// SIMATIC S7-200 project (STEP 7-Micro/WIN), CPU 224 CN REL 02.01

SYMBOL_TABLE Usuario 1
Run              M10.0
Sensor_base      I0.0
X_limite_adelante I0.1
X_limite_atras   I0.2
Y_limite_adelante I0.3
Y_limite_atras   I0.4
Switch           I0.5
Reset            I0.6
Start_y_s1       I0.7
Boton_stop_y_s2  I1.0
Boton_s3_derecha I1.1
Boton_s4_adelante I1.2
Boton_s5_atras   I1.3
Boton_s6_arriba  I1.4
Boton_s7_abajo   I1.5
Pulso_en_Z       Q0.0
Pulso_en_XY      Q0.1
Dir_Eje_Z        Q0.2
Dir_eje_X        Q0.3
Dir_Eje_Y        Q0.4
Pulso_en_X       Q0.5
Pulso_en_Y       Q0.6
Pinza            Q0.7
Posicion_de_Z    VD210
Posicion_de_XY   VD220
Posicion_de_X    VD230
Posicion_de_Y    VD240
Velocidad_de_Z   VD250
Velocidad_de_XY  VD260
END_SYMBOL_TABLE

ORGANIZATION_BLOCK Principal:OB1
TITLE=Notas del programa
BEGIN
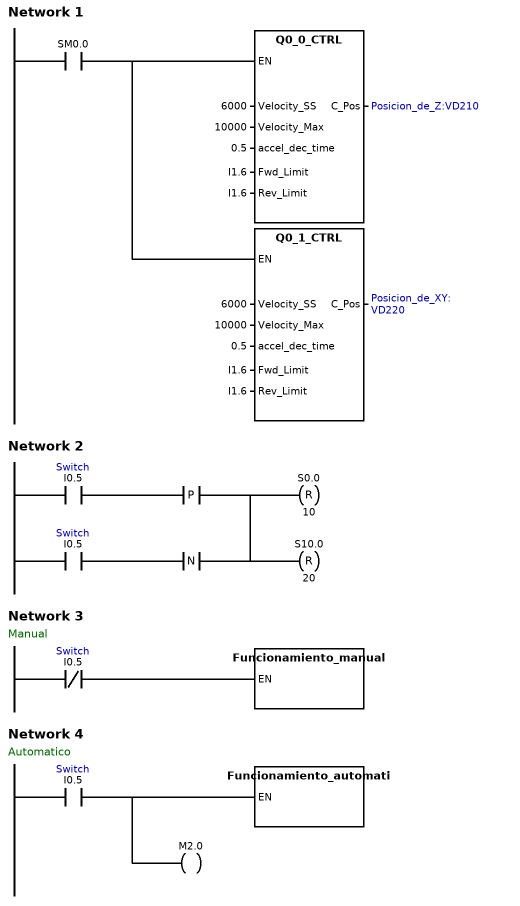
Network 1
// (network saved uncompiled; LAD cells follow)
// row 0: c0 -| |- SM0.0 v  c1 --  c2 [Q0_0_CTRL EN:=power@row0, Velocity_SS:=6000, Velocity_Max:=10000, accel_dec_time:=0.5, Fwd_Limit:=I1.6, Rev_Limit:=I1.6, C_Pos=>Posicion_de_Z:VD210]
// row 1: c0 ^v  c2 [box]
// row 2: c0 ^v  c2 [box]
// row 3: c0 ^  c1 --  c2 [Q0_1_CTRL EN:=power@row3, Velocity_SS:=6000, Velocity_Max:=10000, accel_dec_time:=0.5, Fwd_Limit:=I1.6, Rev_Limit:=I1.6, C_Pos=>Posicion_de_XY:VD220]
// row 4: c2 [box]
// row 5: c2 [box]
Network 2
// (network saved uncompiled; LAD cells follow)
// row 0: c0 -| |- Switch:I0.5  c1 -|P|-  v  c2 -(R) S0.0, 10
// row 1: c0 -| |- Switch:I0.5  c1 -|N|-  ^  c2 -(R) S10.0, 20
Network 3
// Manual
// (network saved uncompiled; LAD cells follow)
// row 0: c0 -|/|- Switch:I0.5  c1 --  c2 [Funcionamiento_manual EN:=power@row0]
Network 4
// Automatico
// (network saved uncompiled; LAD cells follow)
// row 0: c0 -| |- Switch:I0.5 v  c1 --  c2 [Funcionamiento_automati EN:=power@row0]
// row 1: c0 ^  c1 -( ) M2.0
END_ORGANIZATION_BLOCK

SUBROUTINE_BLOCK Funcionamiento_manual:SBR0
TITLE=
BEGIN
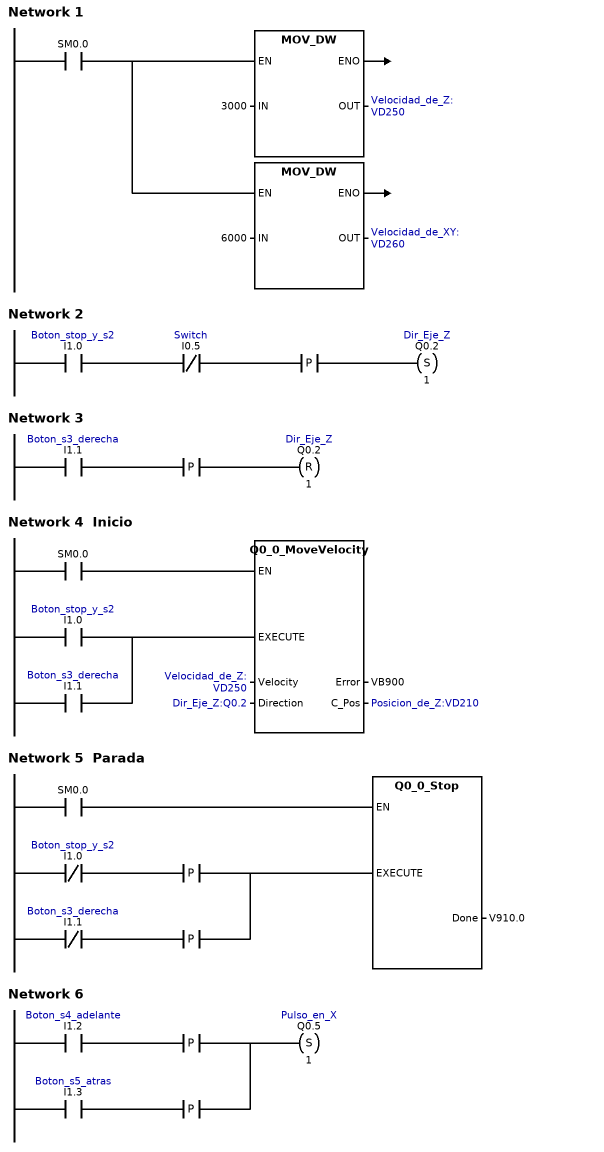
Network 1
// (network saved uncompiled; LAD cells follow)
// row 0: c0 -| |- SM0.0 v  c1 --  c2 [MOV_DW EN:=power@row0, IN:=3000, ENO=>power, OUT=>Velocidad_de_Z:VD250]  c3 ->
// row 1: c0 ^v  c2 [box]
// row 2: c0 ^  c1 --  c2 [MOV_DW EN:=power@row2, IN:=6000, ENO=>power, OUT=>Velocidad_de_XY:VD260]  c3 ->
// row 3: c2 [box]
Network 2
// (network saved uncompiled; LAD cells follow)
// row 0: c0 -| |- Boton_stop_y_s2:I1.0  c1 -|/|- Switch:I0.5  c2 -|P|-  c3 -(S) Dir_Eje_Z:Q0.2, 1
Network 3
// (network saved uncompiled; LAD cells follow)
// row 0: c0 -| |- Boton_s3_derecha:I1.1  c1 -|P|-  c2 -(R) Dir_Eje_Z:Q0.2, 1
Network 4 // Inicio
// (network saved uncompiled; LAD cells follow)
// row 0: c0 -| |- SM0.0  c1 --  c2 [Q0_0_MoveVelocity EN:=power@row0, EXECUTE:=power@row1, Velocity:=Velocidad_de_Z:VD250, Direction:=Dir_Eje_Z:Q0.2, Error=>VB900, C_Pos=>Posicion_de_Z:VD210]
// row 1: c0 -| |- Boton_stop_y_s2:I1.0 v  c1 --  c2 [box]
// row 2: c0 -| |- Boton_s3_derecha:I1.1 ^  c2 [box]
Network 5 // Parada
// (network saved uncompiled; LAD cells follow)
// row 0: c0 -| |- SM0.0  c1 --  c2 --  c3 [Q0_0_Stop EN:=power@row0, EXECUTE:=power@row1, Done=>V910.0]
// row 1: c0 -|/|- Boton_stop_y_s2:I1.0  c1 -|P|-  v  c2 --  c3 [box]
// row 2: c0 -|/|- Boton_s3_derecha:I1.1  c1 -|P|-  ^  c3 [box]
Network 6
// (network saved uncompiled; LAD cells follow)
// row 0: c0 -| |- Boton_s4_adelante:I1.2  c1 -|P|-  v  c2 -(S) Pulso_en_X:Q0.5, 1
// row 1: c0 -| |- Boton_s5_atras:I1.3  c1 -|P|-  ^
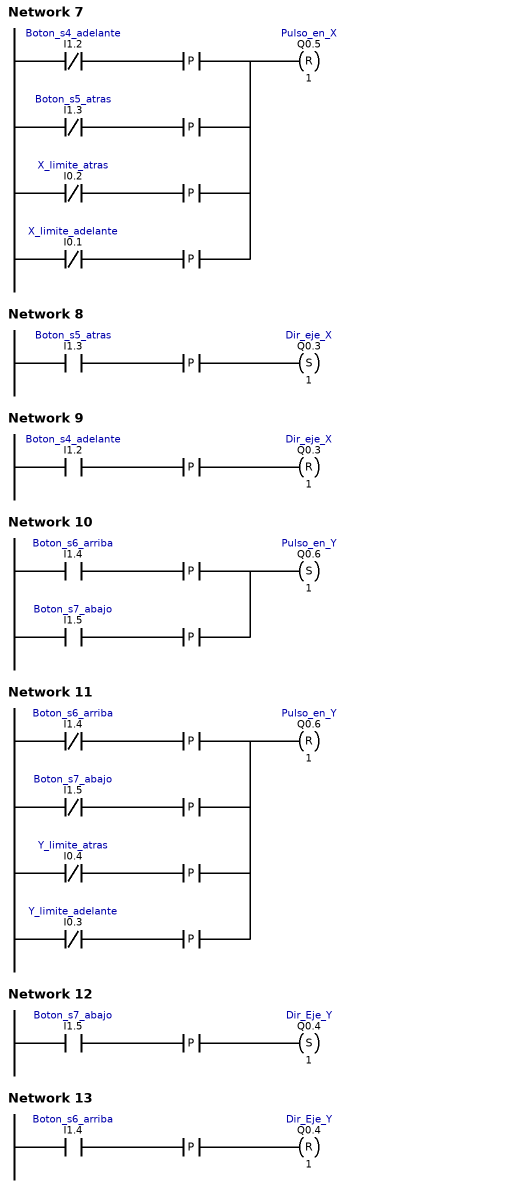
Network 7
// (network saved uncompiled; LAD cells follow)
// row 0: c0 -|/|- Boton_s4_adelante:I1.2  c1 -|P|-  v  c2 -(R) Pulso_en_X:Q0.5, 1
// row 1: c0 -|/|- Boton_s5_atras:I1.3  c1 -|P|-  ^v
// row 2: c0 -|/|- X_limite_atras:I0.2  c1 -|P|-  ^v
// row 3: c0 -|/|- X_limite_adelante:I0.1  c1 -|P|-  ^
Network 8
// (network saved uncompiled; LAD cells follow)
// row 0: c0 -| |- Boton_s5_atras:I1.3  c1 -|P|-  c2 -(S) Dir_eje_X:Q0.3, 1
Network 9
// (network saved uncompiled; LAD cells follow)
// row 0: c0 -| |- Boton_s4_adelante:I1.2  c1 -|P|-  c2 -(R) Dir_eje_X:Q0.3, 1
Network 10
// (network saved uncompiled; LAD cells follow)
// row 0: c0 -| |- Boton_s6_arriba:I1.4  c1 -|P|-  v  c2 -(S) Pulso_en_Y:Q0.6, 1
// row 1: c0 -| |- Boton_s7_abajo:I1.5  c1 -|P|-  ^
Network 11
// (network saved uncompiled; LAD cells follow)
// row 0: c0 -|/|- Boton_s6_arriba:I1.4  c1 -|P|-  v  c2 -(R) Pulso_en_Y:Q0.6, 1
// row 1: c0 -|/|- Boton_s7_abajo:I1.5  c1 -|P|-  ^v
// row 2: c0 -|/|- Y_limite_atras:I0.4  c1 -|P|-  ^v
// row 3: c0 -|/|- Y_limite_adelante:I0.3  c1 -|P|-  ^
Network 12
// (network saved uncompiled; LAD cells follow)
// row 0: c0 -| |- Boton_s7_abajo:I1.5  c1 -|P|-  c2 -(S) Dir_Eje_Y:Q0.4, 1
Network 13
// (network saved uncompiled; LAD cells follow)
// row 0: c0 -| |- Boton_s6_arriba:I1.4  c1 -|P|-  c2 -(R) Dir_Eje_Y:Q0.4, 1
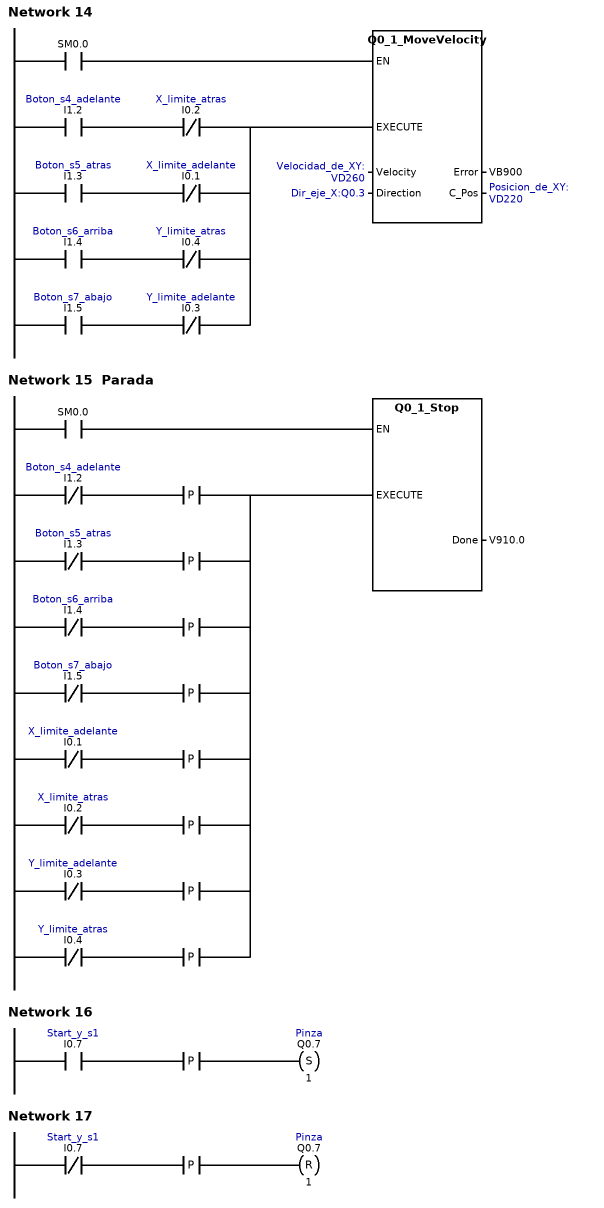
Network 14
// (network saved uncompiled; LAD cells follow)
// row 0: c0 -| |- SM0.0  c1 --  c2 --  c3 [Q0_1_MoveVelocity EN:=power@row0, EXECUTE:=power@row1, Velocity:=Velocidad_de_XY:VD260, Direction:=Dir_eje_X:Q0.3, Error=>VB900, C_Pos=>Posicion_de_XY:VD220]
// row 1: c0 -| |- Boton_s4_adelante:I1.2  c1 -|/|- X_limite_atras:I0.2 v  c2 --  c3 [box]
// row 2: c0 -| |- Boton_s5_atras:I1.3  c1 -|/|- X_limite_adelante:I0.1 ^v  c3 [box]
// row 3: c0 -| |- Boton_s6_arriba:I1.4  c1 -|/|- Y_limite_atras:I0.4 ^v
// row 4: c0 -| |- Boton_s7_abajo:I1.5  c1 -|/|- Y_limite_adelante:I0.3 ^
Network 15 // Parada
// (network saved uncompiled; LAD cells follow)
// row 0: c0 -| |- SM0.0  c1 --  c2 --  c3 [Q0_1_Stop EN:=power@row0, EXECUTE:=power@row1, Done=>V910.0]
// row 1: c0 -|/|- Boton_s4_adelante:I1.2  c1 -|P|-  v  c2 --  c3 [box]
// row 2: c0 -|/|- Boton_s5_atras:I1.3  c1 -|P|-  ^v  c3 [box]
// row 3: c0 -|/|- Boton_s6_arriba:I1.4  c1 -|P|-  ^v
// row 4: c0 -|/|- Boton_s7_abajo:I1.5  c1 -|P|-  ^v
// row 5: c0 -|/|- X_limite_adelante:I0.1  c1 -|P|-  ^v
// row 6: c0 -|/|- X_limite_atras:I0.2  c1 -|P|-  ^v
// row 7: c0 -|/|- Y_limite_adelante:I0.3  c1 -|P|-  ^v
// row 8: c0 -|/|- Y_limite_atras:I0.4  c1 -|P|-  ^
Network 16
// (network saved uncompiled; LAD cells follow)
// row 0: c0 -| |- Start_y_s1:I0.7  c1 -|P|-  c2 -(S) Pinza:Q0.7, 1
Network 17
// (network saved uncompiled; LAD cells follow)
// row 0: c0 -|/|- Start_y_s1:I0.7  c1 -|P|-  c2 -(R) Pinza:Q0.7, 1
Network 22 // 网络标题
// 网络注释
END_SUBROUTINE_BLOCK

// SBR1: protected block, not included

// SBR2: protected block, not included

// SBR3: protected block, not included

// SBR4: protected block, not included

// SBR5: protected block, not included

// SBR6: protected block, not included

SUBROUTINE_BLOCK Origen:SBR7
TITLE=
VAR_INPUT
EXECUTE:BOOL;	// L0.0 
END_VAR
VAR_OUTPUT
Done:BOOL;	// L0.1 
END_VAR
BEGIN
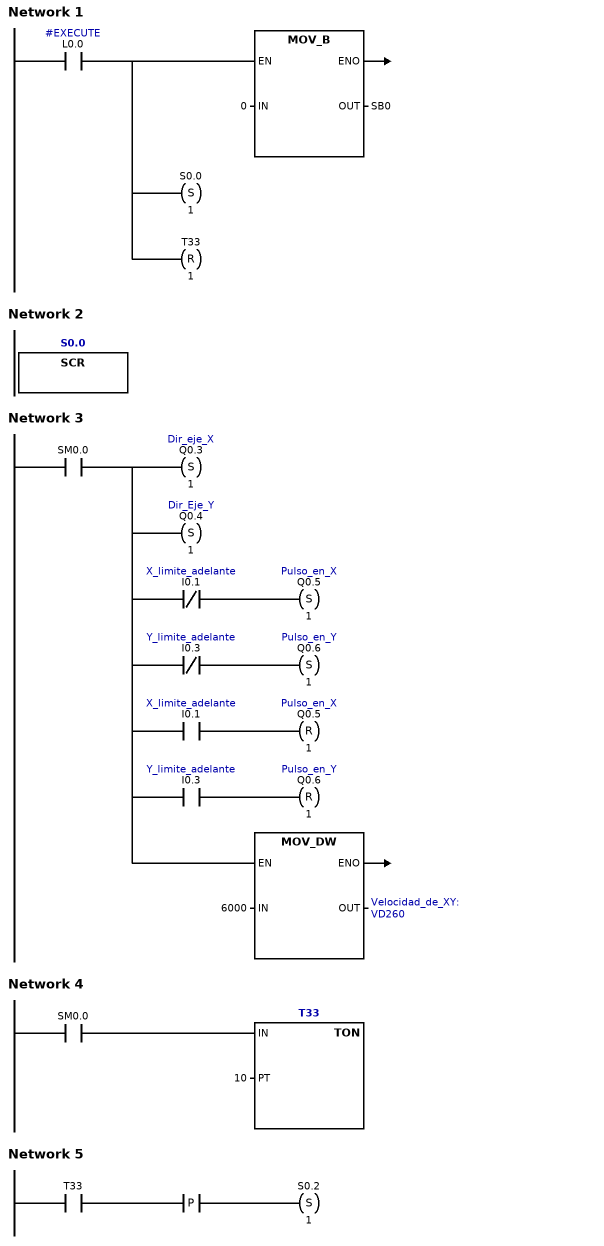
Network 1
LD     #EXECUTE:L0.0
MOVB   0, SB0
S      S0.0, 1
R      T33, 1
Network 2
LSCR   S0.0
Network 3
// (network saved uncompiled; LAD cells follow)
// row 0: c0 -| |- SM0.0 v  c1 -(S) Dir_eje_X:Q0.3, 1
// row 1: c0 ^v  c1 -(S) Dir_Eje_Y:Q0.4, 1
// row 2: c0 ^v  c1 -|/|- X_limite_adelante:I0.1  c2 -(S) Pulso_en_X:Q0.5, 1
// row 3: c0 ^v  c1 -|/|- Y_limite_adelante:I0.3  c2 -(S) Pulso_en_Y:Q0.6, 1
// row 4: c0 ^v  c1 -| |- X_limite_adelante:I0.1  c2 -(R) Pulso_en_X:Q0.5, 1
// row 5: c0 ^v  c1 -| |- Y_limite_adelante:I0.3  c2 -(R) Pulso_en_Y:Q0.6, 1
// row 6: c0 ^  c1 --  c2 [MOV_DW EN:=power@row6, IN:=6000, ENO=>power, OUT=>Velocidad_de_XY:VD260]  c3 ->
// row 7: c2 [box]
Network 4
LD     SM0.0
TON    T33, 10
Network 5
LD     T33
EU
S      S0.2, 1
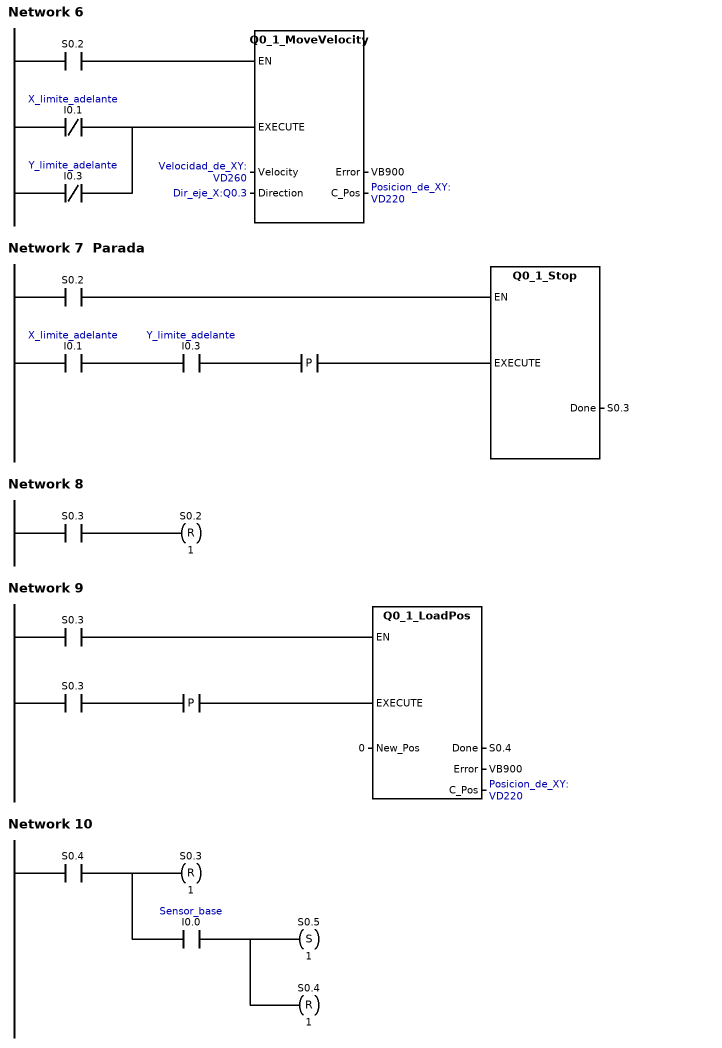
Network 6
// (network saved uncompiled; LAD cells follow)
// row 0: c0 -| |- S0.2  c1 --  c2 [Q0_1_MoveVelocity EN:=power@row0, EXECUTE:=power@row1, Velocity:=Velocidad_de_XY:VD260, Direction:=Dir_eje_X:Q0.3, Error=>VB900, C_Pos=>Posicion_de_XY:VD220]
// row 1: c0 -|/|- X_limite_adelante:I0.1 v  c1 --  c2 [box]
// row 2: c0 -|/|- Y_limite_adelante:I0.3 ^  c2 [box]
Network 7 // Parada
// (network saved uncompiled; LAD cells follow)
// row 0: c0 -| |- S0.2  c1 --  c2 --  c3 --  c4 [Q0_1_Stop EN:=power@row0, EXECUTE:=power@row1, Done=>S0.3]
// row 1: c0 -| |- X_limite_adelante:I0.1  c1 -| |- Y_limite_adelante:I0.3  c2 -|P|-  c3 --  c4 [box]
// row 2: c4 [box]
Network 8
LD     S0.3
R      S0.2, 1
Network 9
// (network saved uncompiled; LAD cells follow)
// row 0: c0 -| |- S0.3  c1 --  c2 --  c3 [Q0_1_LoadPos EN:=power@row0, EXECUTE:=power@row1, New_Pos:=0, Done=>S0.4, Error=>VB900, C_Pos=>Posicion_de_XY:VD220]
// row 1: c0 -| |- S0.3  c1 -|P|-  c2 --  c3 [box]
// row 2: c3 [box]
Network 10
// (network saved uncompiled; LAD cells follow)
// row 0: c0 -| |- S0.4 v  c1 -(R) S0.3, 1
// row 1: c0 ^  c1 -| |- Sensor_base:I0.0 v  c2 -(S) S0.5, 1
// row 2: c1 ^  c2 -(R) S0.4, 1
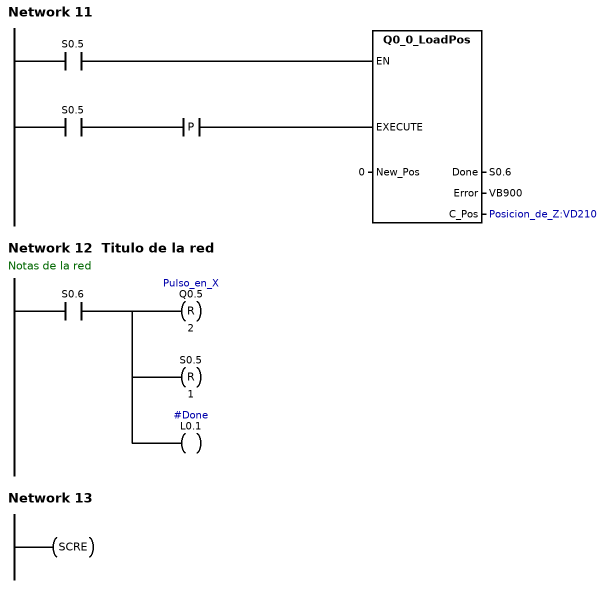
Network 11
// (network saved uncompiled; LAD cells follow)
// row 0: c0 -| |- S0.5  c1 --  c2 --  c3 [Q0_0_LoadPos EN:=power@row0, EXECUTE:=power@row1, New_Pos:=0, Done=>S0.6, Error=>VB900, C_Pos=>Posicion_de_Z:VD210]
// row 1: c0 -| |- S0.5  c1 -|P|-  c2 --  c3 [box]
// row 2: c3 [box]
Network 12 // Titulo de la red
// Notas de la red
// (network saved uncompiled; LAD cells follow)
// row 0: c0 -| |- S0.6 v  c1 -(R) Pulso_en_X:Q0.5, 2
// row 1: c0 ^v  c1 -(R) S0.5, 1
// row 2: c0 ^  c1 -( ) #Done:L0.1
Network 13
SCRE
Network 25 // 网络标题
// 网络注释
END_SUBROUTINE_BLOCK

SUBROUTINE_BLOCK Funcionamiento_automati:SBR8
TITLE=
BEGIN
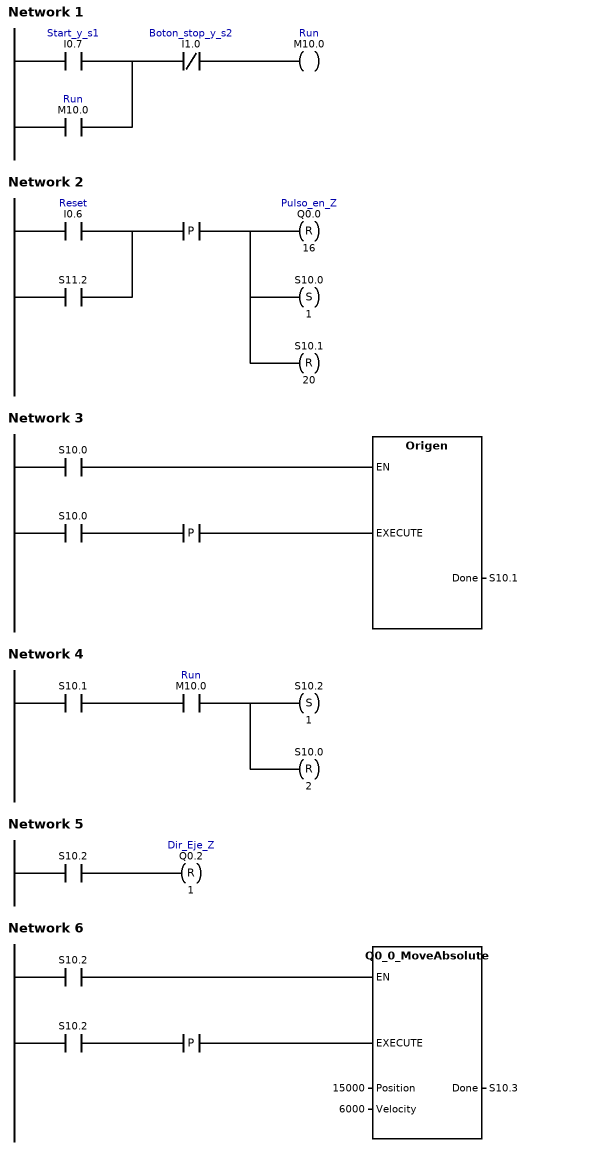
Network 1
// (network saved uncompiled; LAD cells follow)
// row 0: c0 -| |- Start_y_s1:I0.7 v  c1 -|/|- Boton_stop_y_s2:I1.0  c2 -( ) Run:M10.0
// row 1: c0 -| |- Run:M10.0 ^
Network 2
// (network saved uncompiled; LAD cells follow)
// row 0: c0 -| |- Reset:I0.6 v  c1 -|P|-  v  c2 -(R) Pulso_en_Z:Q0.0, 16
// row 1: c0 -| |- S11.2 ^  c1 ^v  c2 -(S) S10.0, 1
// row 2: c1 ^  c2 -(R) S10.1, 20
Network 3
LD     S10.0
=      L60.0
LD     S10.0
EU
=      L63.7
LD     L60.0
CALL   Origen:SBR7, L63.7, S10.1
Network 4
// (network saved uncompiled; LAD cells follow)
// row 0: c0 -| |- S10.1  c1 -| |- Run:M10.0 v  c2 -(S) S10.2, 1
// row 1: c1 ^  c2 -(R) S10.0, 2
Network 5
// (network saved uncompiled; LAD cells follow)
// row 0: c0 -| |- S10.2  c1 -(R) Dir_Eje_Z:Q0.2, 1
Network 6
LD     S10.2
=      L60.0
LD     S10.2
EU
=      L63.7
LD     L60.0
CALL   Q0_0_MoveAbsolute:SBR4, L63.7, 15000, 6000, S10.3
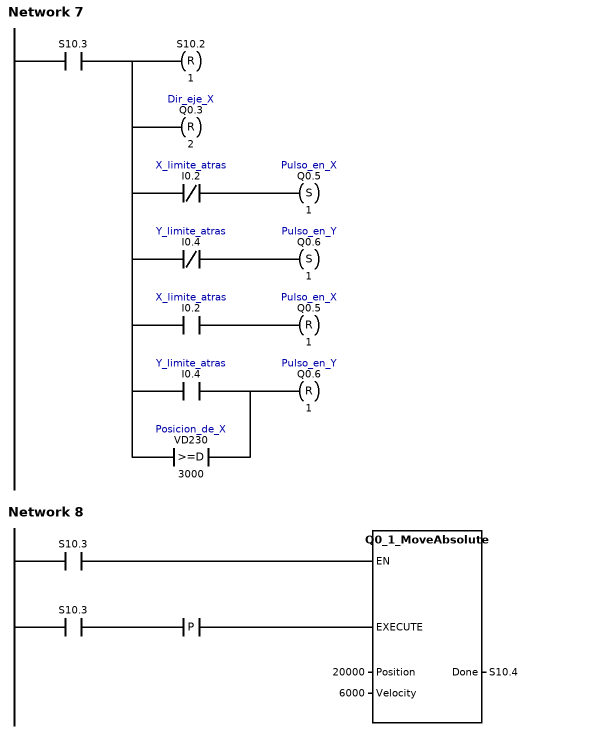
Network 7
// (network saved uncompiled; LAD cells follow)
// row 0: c0 -| |- S10.3 v  c1 -(R) S10.2, 1
// row 1: c0 ^v  c1 -(R) Dir_eje_X:Q0.3, 2
// row 2: c0 ^v  c1 -|/|- X_limite_atras:I0.2  c2 -(S) Pulso_en_X:Q0.5, 1
// row 3: c0 ^v  c1 -|/|- Y_limite_atras:I0.4  c2 -(S) Pulso_en_Y:Q0.6, 1
// row 4: c0 ^v  c1 -| |- X_limite_atras:I0.2  c2 -(R) Pulso_en_X:Q0.5, 1
// row 5: c0 ^v  c1 -| |- Y_limite_atras:I0.4 v  c2 -(R) Pulso_en_Y:Q0.6, 1
// row 6: c0 ^  c1 -|>=D|- Posicion_de_X:VD230, 3000 ^
Network 8
LD     S10.3
=      L60.0
LD     S10.3
EU
=      L63.7
LD     L60.0
CALL   Q0_1_MoveAbsolute:SBR19, L63.7, 20000, 6000, S10.4
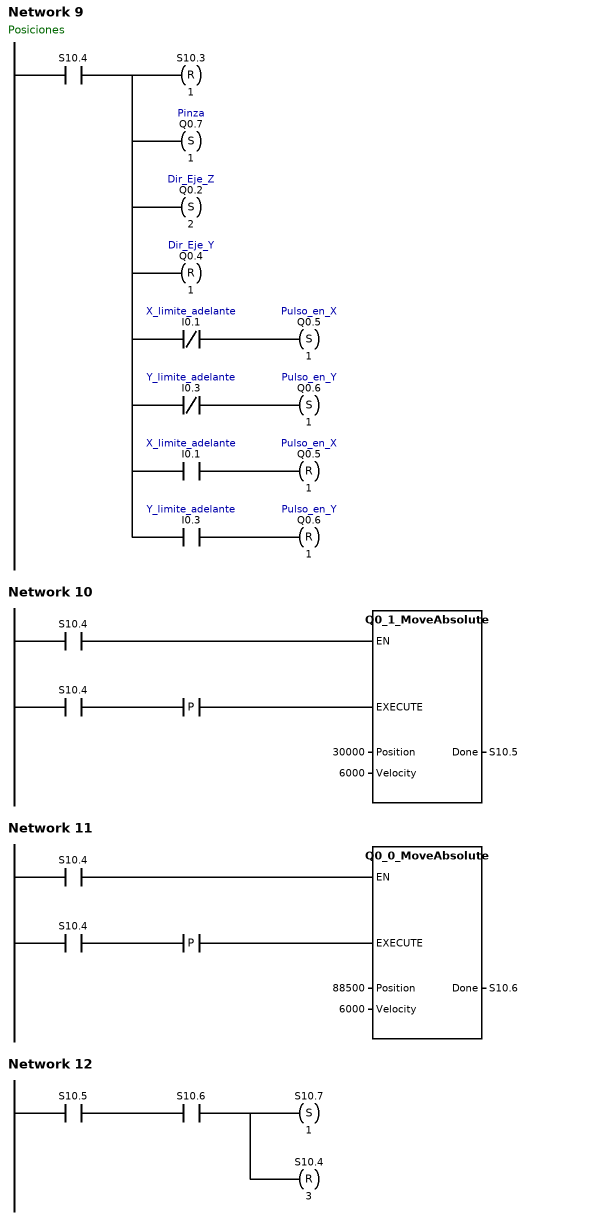
Network 9
// Posiciones
// (network saved uncompiled; LAD cells follow)
// row 0: c0 -| |- S10.4 v  c1 -(R) S10.3, 1
// row 1: c0 ^v  c1 -(S) Pinza:Q0.7, 1
// row 2: c0 ^v  c1 -(S) Dir_Eje_Z:Q0.2, 2
// row 3: c0 ^v  c1 -(R) Dir_Eje_Y:Q0.4, 1
// row 4: c0 ^v  c1 -|/|- X_limite_adelante:I0.1  c2 -(S) Pulso_en_X:Q0.5, 1
// row 5: c0 ^v  c1 -|/|- Y_limite_adelante:I0.3  c2 -(S) Pulso_en_Y:Q0.6, 1
// row 6: c0 ^v  c1 -| |- X_limite_adelante:I0.1  c2 -(R) Pulso_en_X:Q0.5, 1
// row 7: c0 ^  c1 -| |- Y_limite_adelante:I0.3  c2 -(R) Pulso_en_Y:Q0.6, 1
Network 10
LD     S10.4
=      L60.0
LD     S10.4
EU
=      L63.7
LD     L60.0
CALL   Q0_1_MoveAbsolute:SBR19, L63.7, 30000, 6000, S10.5
Network 11
LD     S10.4
=      L60.0
LD     S10.4
EU
=      L63.7
LD     L60.0
CALL   Q0_0_MoveAbsolute:SBR4, L63.7, 88500, 6000, S10.6
Network 12
LD     S10.5
A      S10.6
S      S10.7, 1
R      S10.4, 3
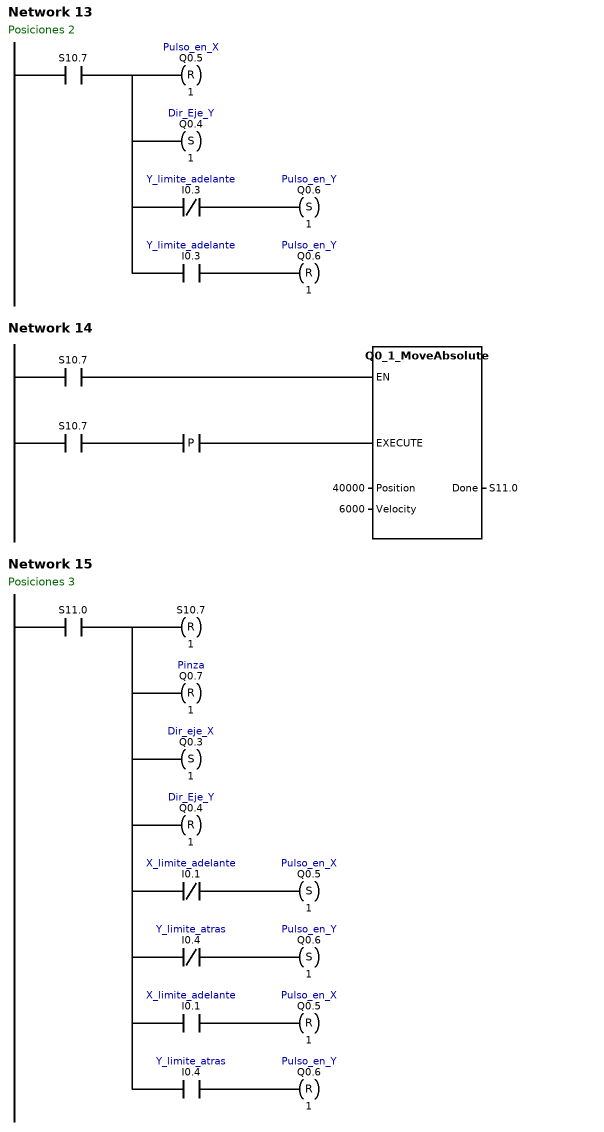
Network 13
// Posiciones 2
// (network saved uncompiled; LAD cells follow)
// row 0: c0 -| |- S10.7 v  c1 -(R) Pulso_en_X:Q0.5, 1
// row 1: c0 ^v  c1 -(S) Dir_Eje_Y:Q0.4, 1
// row 2: c0 ^v  c1 -|/|- Y_limite_adelante:I0.3  c2 -(S) Pulso_en_Y:Q0.6, 1
// row 3: c0 ^  c1 -| |- Y_limite_adelante:I0.3  c2 -(R) Pulso_en_Y:Q0.6, 1
Network 14
LD     S10.7
=      L60.0
LD     S10.7
EU
=      L63.7
LD     L60.0
CALL   Q0_1_MoveAbsolute:SBR19, L63.7, 40000, 6000, S11.0
Network 15
// Posiciones 3
// (network saved uncompiled; LAD cells follow)
// row 0: c0 -| |- S11.0 v  c1 -(R) S10.7, 1
// row 1: c0 ^v  c1 -(R) Pinza:Q0.7, 1
// row 2: c0 ^v  c1 -(S) Dir_eje_X:Q0.3, 1
// row 3: c0 ^v  c1 -(R) Dir_Eje_Y:Q0.4, 1
// row 4: c0 ^v  c1 -|/|- X_limite_adelante:I0.1  c2 -(S) Pulso_en_X:Q0.5, 1
// row 5: c0 ^v  c1 -|/|- Y_limite_atras:I0.4  c2 -(S) Pulso_en_Y:Q0.6, 1
// row 6: c0 ^v  c1 -| |- X_limite_adelante:I0.1  c2 -(R) Pulso_en_X:Q0.5, 1
// row 7: c0 ^  c1 -| |- Y_limite_atras:I0.4  c2 -(R) Pulso_en_Y:Q0.6, 1
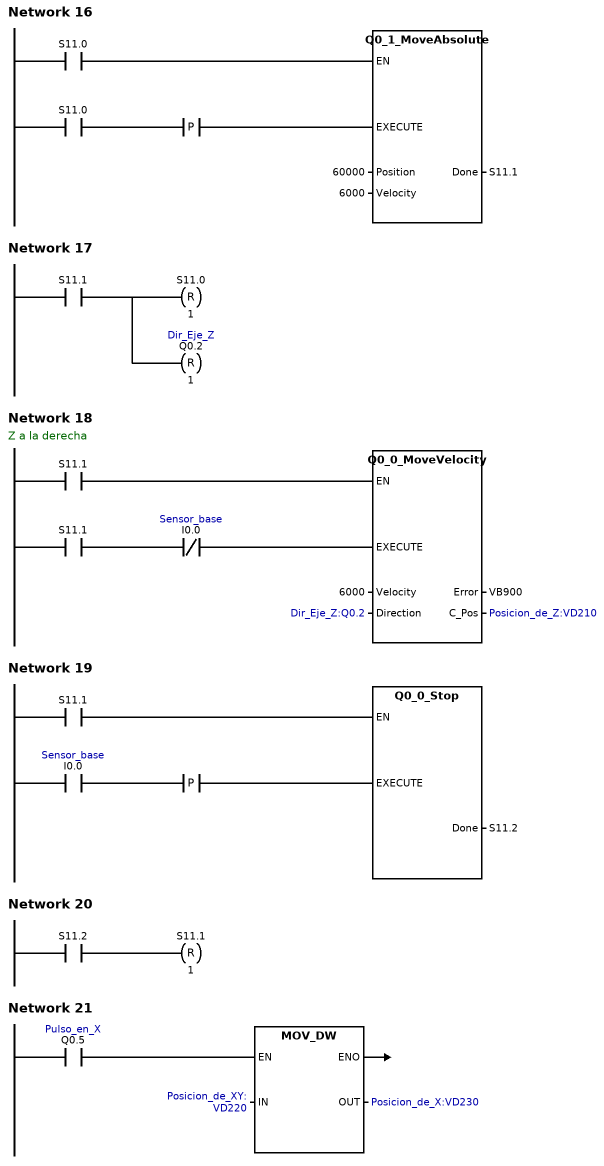
Network 16
LD     S11.0
=      L60.0
LD     S11.0
EU
=      L63.7
LD     L60.0
CALL   Q0_1_MoveAbsolute:SBR19, L63.7, 60000, 6000, S11.1
Network 17
// (network saved uncompiled; LAD cells follow)
// row 0: c0 -| |- S11.1 v  c1 -(R) S11.0, 1
// row 1: c0 ^  c1 -(R) Dir_Eje_Z:Q0.2, 1
Network 18
// Z a la derecha
// (network saved uncompiled; LAD cells follow)
// row 0: c0 -| |- S11.1  c1 --  c2 --  c3 [Q0_0_MoveVelocity EN:=power@row0, EXECUTE:=power@row1, Velocity:=6000, Direction:=Dir_Eje_Z:Q0.2, Error=>VB900, C_Pos=>Posicion_de_Z:VD210]
// row 1: c0 -| |- S11.1  c1 -|/|- Sensor_base:I0.0  c2 --  c3 [box]
// row 2: c3 [box]
Network 19
// (network saved uncompiled; LAD cells follow)
// row 0: c0 -| |- S11.1  c1 --  c2 --  c3 [Q0_0_Stop EN:=power@row0, EXECUTE:=power@row1, Done=>S11.2]
// row 1: c0 -| |- Sensor_base:I0.0  c1 -|P|-  c2 --  c3 [box]
// row 2: c3 [box]
Network 20
LD     S11.2
R      S11.1, 1
Network 21
// (network saved uncompiled; LAD cells follow)
// row 0: c0 -| |- Pulso_en_X:Q0.5  c1 --  c2 [MOV_DW EN:=power@row0, IN:=Posicion_de_XY:VD220, ENO=>power, OUT=>Posicion_de_X:VD230]  c3 ->
// row 1: c2 [box]
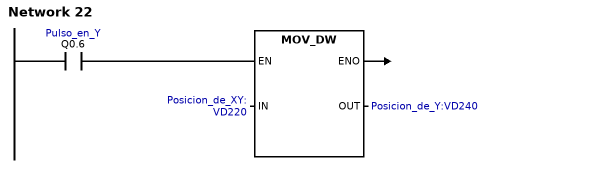
Network 22
// (network saved uncompiled; LAD cells follow)
// row 0: c0 -| |- Pulso_en_Y:Q0.6  c1 --  c2 [MOV_DW EN:=power@row0, IN:=Posicion_de_XY:VD220, ENO=>power, OUT=>Posicion_de_Y:VD240]  c3 ->
// row 1: c2 [box]
END_SUBROUTINE_BLOCK

// SBR9: protected block, not included

// SBR10: protected block, not included

// SBR11: protected block, not included

// SBR12: protected block, not included

// SBR13: protected block, not included

// SBR14: protected block, not included

// SBR15: protected block, not included

// SBR16: protected block, not included

// SBR17: protected block, not included

// SBR18: protected block, not included
